FUNCTION_BLOCK logiBUS_QD_SDM_G (* Output service interface function block for a sigma-delta output with gamma correction for LEDs (brightness 0..8191 in DWORD, 8 bit pulse density, 1 MHz). Logic level only: LEDs, LED drivers, not the power outputs *)
  (* Standard: 61499-2; Description: Copyright (c) 2026 HR Agrartechnik GmbH This program and the accompanying materials are made available under the terms of the Eclipse Public License 2.0 which is available at https://www.eclipse.org/legal/epl-2.0/ SPDX-License-Identifier: EPL-2.0 *)
  (* Version 1.0, 2026-11-06, Franz Höpfinger, HR Agrartechnik GmbH, initial version *)
  PACKAGE logiBUS::io::DQ;
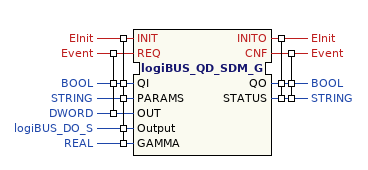
  EVENT_INPUT
    INIT : EInit WITH QI, PARAMS, Output, GAMMA; (* Service Initialization *)
    REQ WITH QI, OUT; (* Service Request *)
  END_EVENT
  EVENT_OUTPUT
    INITO : EInit WITH QO, STATUS; (* Initialization Confirm *)
    CNF WITH QO, STATUS; (* Confirmation of Requested Service *)
  END_EVENT
  VAR_INPUT
    QI : BOOL; (* Event Input Qualifier *)
    PARAMS : STRING; (* Service Parameters *)
    OUT : DWORD; (* Brightness as the eye sees it (0..8191), converted with GAMMA, output as pulse density with 8 bit (256 steps). No ramp *)
    Output : logiBUS::io::DQ::logiBUS_DO_S := logiBUS_DO::Invalid; (* Identify the Output Output_Q1..Q8 *)
    GAMMA : REAL := 2.2; (* Gamma of the brightness curve, read at INIT: density from (OUT / 8191)^GAMMA. 1.0 = linear, 2.2 = sRGB (default). Invalid values (<= 0, not finite) run linear like 1.0. With 8 bit the lowest steps become coarse *)
  END_VAR
  VAR_OUTPUT
    QO : BOOL; (* Event Output Qualifier *)
    STATUS : STRING; (* Service Status *)
  END_VAR
END_FUNCTION_BLOCK
